// Vérifier, activer ou annuler la zone d'attente (docs/05 § 10)
{attribute 'pack_mode' := '1'}
TYPE ST_DeployRequest :
STRUCT
    nSeq : UDINT;
    eCmd : E_DeployCmd;
    nCrcMachine : UDINT;
    aCrcStation : ARRAY[1..GVL_Const.MAX_STATIONS] OF UDINT;
    nCrcRecipes : UDINT;
    nInstrSetRequired : UINT;       // docs/02 § 7.3
    nCatalogRequired : UINT;
    sUser : STRING(24);
END_STRUCT
END_TYPE

(* stored: Version 1.1.0.1, ProductVersion 3.1.4024.12
   DUT ST_DeployRequest: Id {55a1a67f-9ded-513d-bbdc-b6a426112c2b} *)
